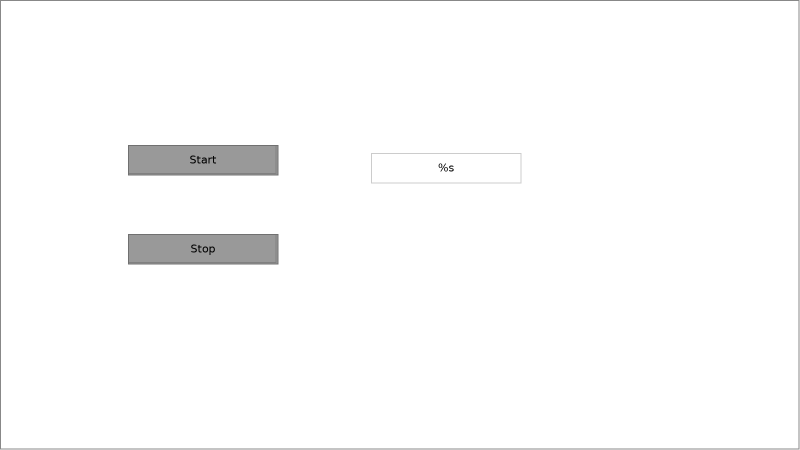
VISUALIZATION Main  // 800x450
    Button (128,145 150x30), "Start"
        tap GVL.bStart
    Button (128,234 150x30), "Stop"
        tap GVL.bStop
    Textfield (371,153 150x30), "%s", text variable: MAIN.fbCTU3.CV
END_VISUALIZATION

(* stored: Version 1.1.0.1, ProductVersion 3.1.4026.18
   Visu Main: Id {d2832147-dbf0-4274-9036-5216bbb99c82} *)
